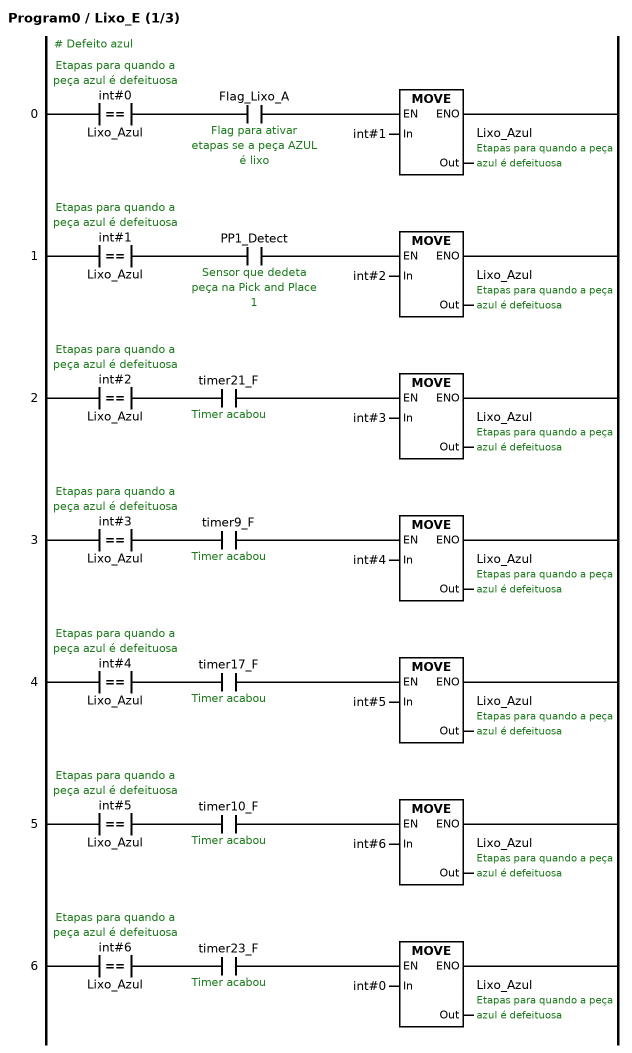
(* [picture p120: Program0 / Lixo_E, rungs 0-6] *)
(* Rung 0: # Defeito azul *)
IF (int#0 = Lixo_Azul) AND Flag_Lixo_A THEN Lixo_Azul := int#1; END_IF;
(* Rung 1 *)
IF (int#1 = Lixo_Azul) AND PP1_Detect THEN Lixo_Azul := int#2; END_IF;
(* Rung 2 *)
IF (int#2 = Lixo_Azul) AND timer21_F THEN Lixo_Azul := int#3; END_IF;
(* Rung 3 *)
IF (int#3 = Lixo_Azul) AND timer9_F THEN Lixo_Azul := int#4; END_IF;
(* Rung 4 *)
IF (int#4 = Lixo_Azul) AND timer17_F THEN Lixo_Azul := int#5; END_IF;
(* Rung 5 *)
IF (int#5 = Lixo_Azul) AND timer10_F THEN Lixo_Azul := int#6; END_IF;
(* Rung 6 *)
IF (int#6 = Lixo_Azul) AND timer23_F THEN Lixo_Azul := int#0; END_IF;

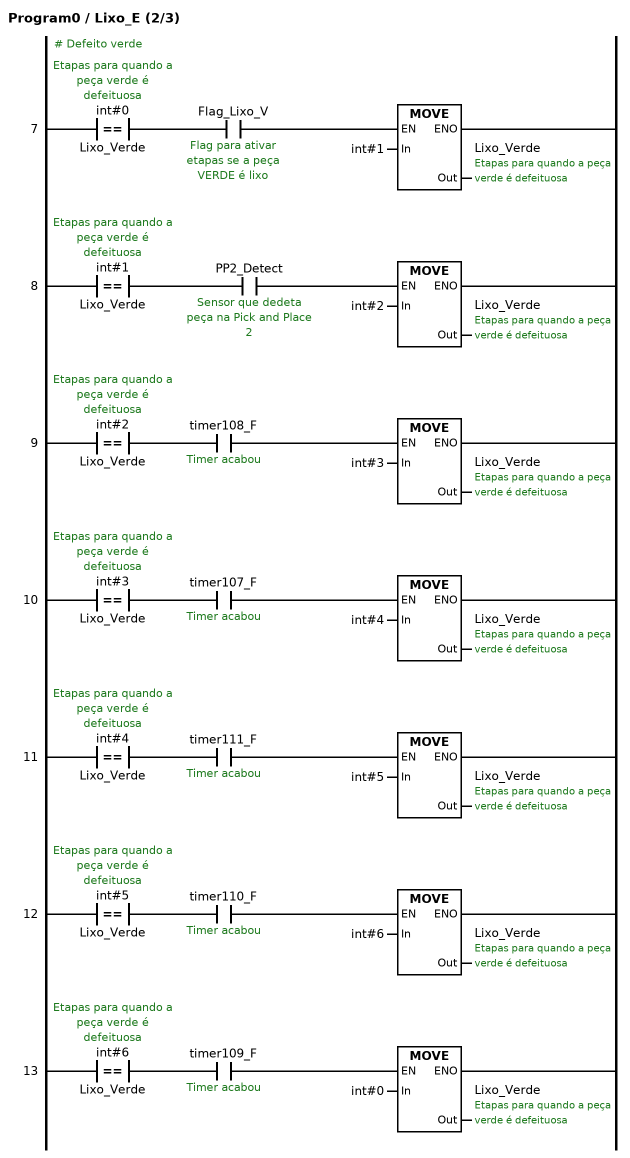
(* Rung 7: # Defeito verde *)
IF (int#0 = Lixo_Verde) AND Flag_Lixo_V THEN Lixo_Verde := int#1; END_IF;
(* Rung 8 *)
IF (int#1 = Lixo_Verde) AND PP2_Detect THEN Lixo_Verde := int#2; END_IF;
(* Rung 9 *)
IF (int#2 = Lixo_Verde) AND timer108_F THEN Lixo_Verde := int#3; END_IF;
(* Rung 10 *)
IF (int#3 = Lixo_Verde) AND timer107_F THEN Lixo_Verde := int#4; END_IF;
(* Rung 11 *)
IF (int#4 = Lixo_Verde) AND timer111_F THEN Lixo_Verde := int#5; END_IF;
(* Rung 12 *)
IF (int#5 = Lixo_Verde) AND timer110_F THEN Lixo_Verde := int#6; END_IF;
(* Rung 13 *)
IF (int#6 = Lixo_Verde) AND timer109_F THEN Lixo_Verde := int#0; END_IF;

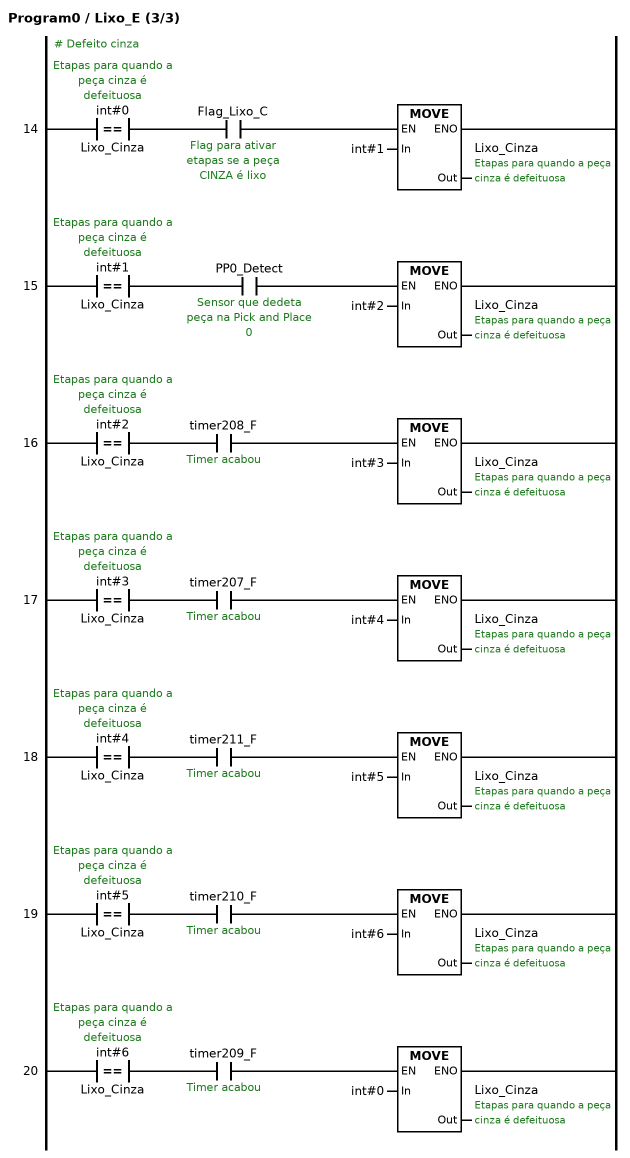
(* Rung 14: # Defeito cinza *)
IF (int#0 = Lixo_Cinza) AND Flag_Lixo_C THEN Lixo_Cinza := int#1; END_IF;
(* Rung 15 *)
IF (int#1 = Lixo_Cinza) AND PP0_Detect THEN Lixo_Cinza := int#2; END_IF;
(* Rung 16 *)
IF (int#2 = Lixo_Cinza) AND timer208_F THEN Lixo_Cinza := int#3; END_IF;
(* Rung 17 *)
IF (int#3 = Lixo_Cinza) AND timer207_F THEN Lixo_Cinza := int#4; END_IF;
(* Rung 18 *)
IF (int#4 = Lixo_Cinza) AND timer211_F THEN Lixo_Cinza := int#5; END_IF;
(* Rung 19 *)
IF (int#5 = Lixo_Cinza) AND timer210_F THEN Lixo_Cinza := int#6; END_IF;
(* Rung 20 *)
IF (int#6 = Lixo_Cinza) AND timer209_F THEN Lixo_Cinza := int#0; END_IF;

(* Section Lixo_S: ladder, written here as Structured Text *)

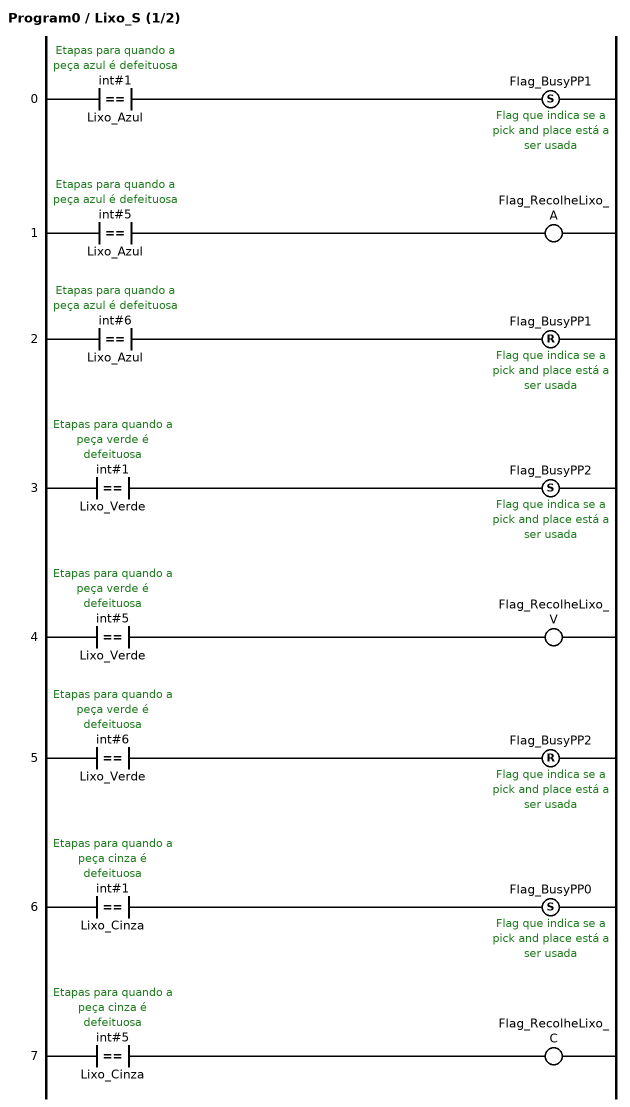
(* Rung 0 *)
IF int#1 = Lixo_Azul THEN Flag_BusyPP1 := TRUE; END_IF;
(* Rung 1 *)
Flag_RecolheLixo_A := int#5 = Lixo_Azul;
(* Rung 2 *)
IF int#6 = Lixo_Azul THEN Flag_BusyPP1 := FALSE; END_IF;
(* Rung 3 *)
IF int#1 = Lixo_Verde THEN Flag_BusyPP2 := TRUE; END_IF;
(* Rung 4 *)
Flag_RecolheLixo_V := int#5 = Lixo_Verde;
(* Rung 5 *)
IF int#6 = Lixo_Verde THEN Flag_BusyPP2 := FALSE; END_IF;
(* Rung 6 *)
IF int#1 = Lixo_Cinza THEN Flag_BusyPP0 := TRUE; END_IF;
(* Rung 7 *)
Flag_RecolheLixo_C := int#5 = Lixo_Cinza;

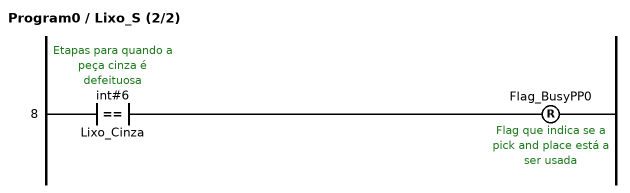
(* Rung 8 *)
IF int#6 = Lixo_Cinza THEN Flag_BusyPP0 := FALSE; END_IF;

(* Section Recolhe_Lixo_E: ladder, written here as Structured Text *)

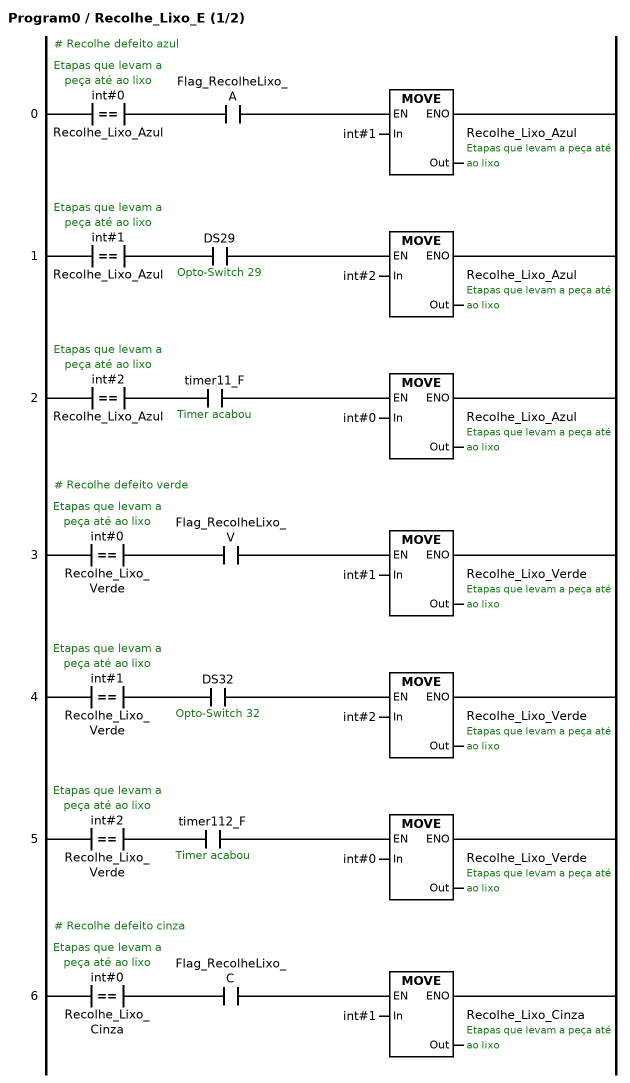
(* Rung 0: # Recolhe defeito azul *)
IF (int#0 = Recolhe_Lixo_Azul) AND Flag_RecolheLixo_A THEN Recolhe_Lixo_Azul := int#1; END_IF;
(* Rung 1 *)
IF (int#1 = Recolhe_Lixo_Azul) AND DS29 THEN Recolhe_Lixo_Azul := int#2; END_IF;
(* Rung 2 *)
IF (int#2 = Recolhe_Lixo_Azul) AND timer11_F THEN Recolhe_Lixo_Azul := int#0; END_IF;
(* Rung 3: # Recolhe defeito verde *)
IF (int#0 = Recolhe_Lixo_Verde) AND Flag_RecolheLixo_V THEN Recolhe_Lixo_Verde := int#1; END_IF;
(* Rung 4 *)
IF (int#1 = Recolhe_Lixo_Verde) AND DS32 THEN Recolhe_Lixo_Verde := int#2; END_IF;
(* Rung 5 *)
IF (int#2 = Recolhe_Lixo_Verde) AND timer112_F THEN Recolhe_Lixo_Verde := int#0; END_IF;
(* Rung 6: # Recolhe defeito cinza *)
IF (int#0 = Recolhe_Lixo_Cinza) AND Flag_RecolheLixo_C THEN Recolhe_Lixo_Cinza := int#1; END_IF;

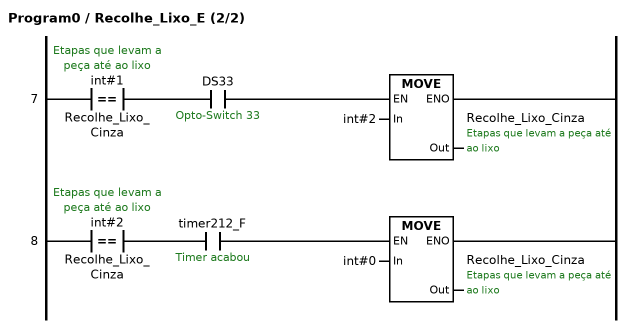
(* Rung 7 *)
IF (int#1 = Recolhe_Lixo_Cinza) AND DS33 THEN Recolhe_Lixo_Cinza := int#2; END_IF;
(* Rung 8 *)
IF (int#2 = Recolhe_Lixo_Cinza) AND timer212_F THEN Recolhe_Lixo_Cinza := int#0; END_IF;

(* Section Recolhe_Lixo_S: ladder, written here as Structured Text *)

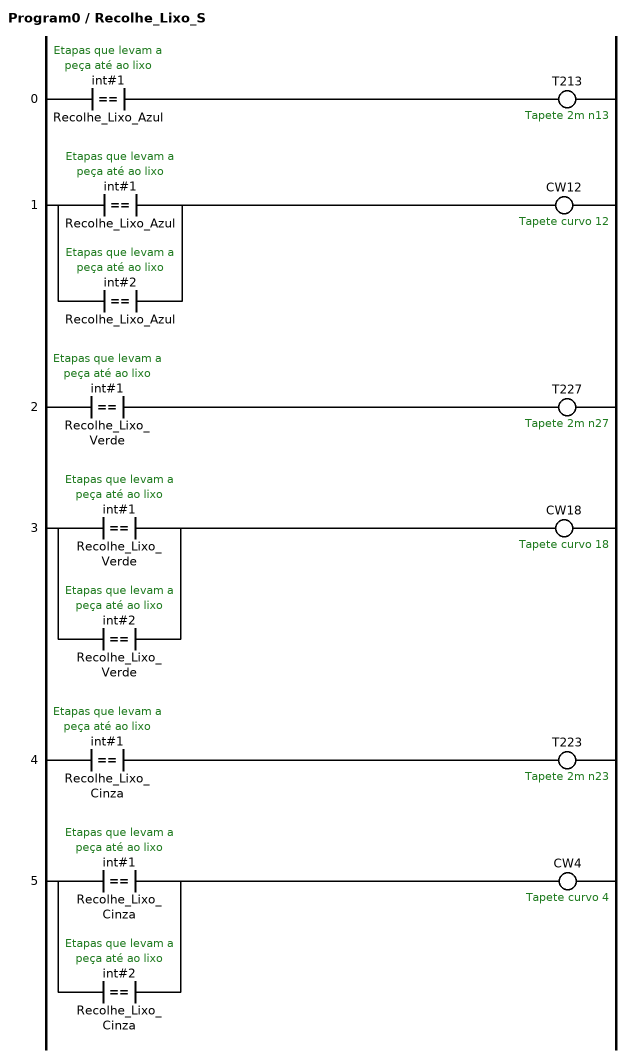
(* Rung 0 *)
T213 := int#1 = Recolhe_Lixo_Azul;
(* Rung 1 *)
CW12 := (int#1 = Recolhe_Lixo_Azul) OR (int#2 = Recolhe_Lixo_Azul);
(* Rung 2 *)
T227 := int#1 = Recolhe_Lixo_Verde;
(* Rung 3 *)
CW18 := (int#1 = Recolhe_Lixo_Verde) OR (int#2 = Recolhe_Lixo_Verde);
(* Rung 4 *)
T223 := int#1 = Recolhe_Lixo_Cinza;
(* Rung 5 *)
CW4 := (int#1 = Recolhe_Lixo_Cinza) OR (int#2 = Recolhe_Lixo_Cinza);

(* Section Repara_Peca_E: ladder, written here as Structured Text *)

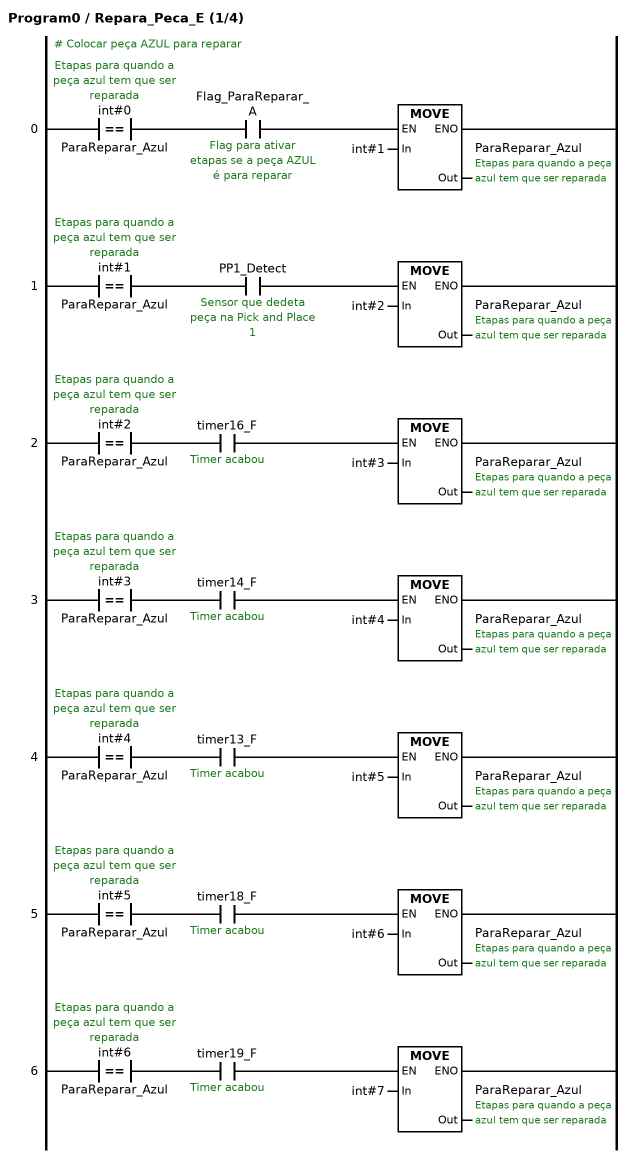
(* Rung 0: # Colocar peça AZUL para reparar *)
IF (int#0 = ParaReparar_Azul) AND Flag_ParaReparar_A THEN ParaReparar_Azul := int#1; END_IF;
(* Rung 1 *)
IF (int#1 = ParaReparar_Azul) AND PP1_Detect THEN ParaReparar_Azul := int#2; END_IF;
(* Rung 2 *)
IF (int#2 = ParaReparar_Azul) AND timer16_F THEN ParaReparar_Azul := int#3; END_IF;
(* Rung 3 *)
IF (int#3 = ParaReparar_Azul) AND timer14_F THEN ParaReparar_Azul := int#4; END_IF;
(* Rung 4 *)
IF (int#4 = ParaReparar_Azul) AND timer13_F THEN ParaReparar_Azul := int#5; END_IF;
(* Rung 5 *)
IF (int#5 = ParaReparar_Azul) AND timer18_F THEN ParaReparar_Azul := int#6; END_IF;
(* Rung 6 *)
IF (int#6 = ParaReparar_Azul) AND timer19_F THEN ParaReparar_Azul := int#7; END_IF;

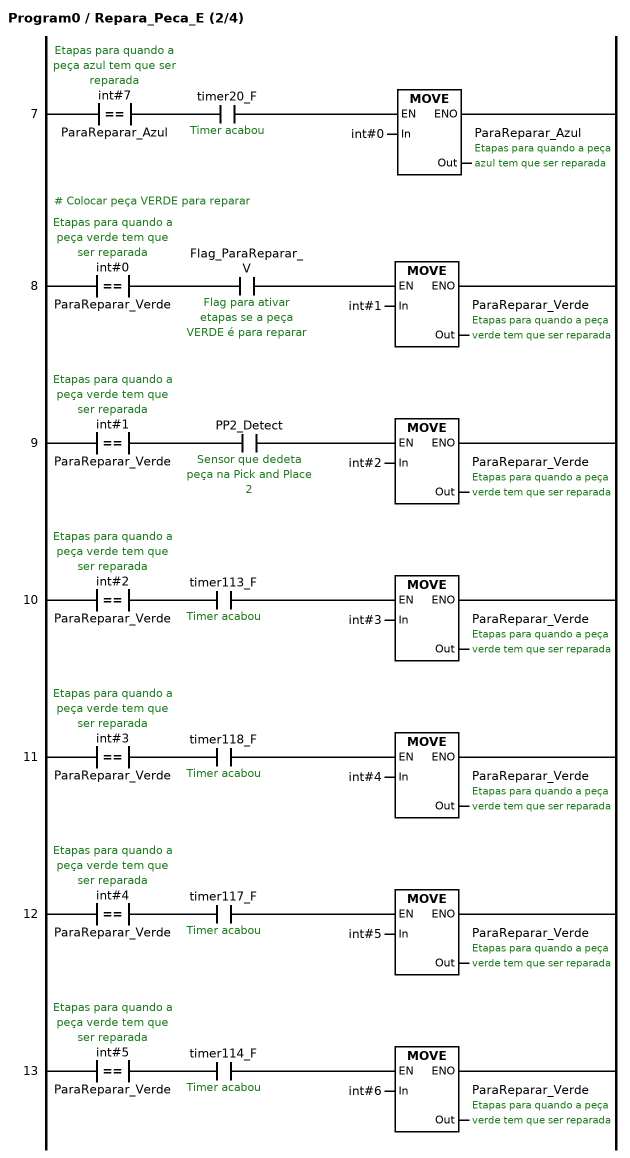
(* Rung 7 *)
IF (int#7 = ParaReparar_Azul) AND timer20_F THEN ParaReparar_Azul := int#0; END_IF;
(* Rung 8: # Colocar peça VERDE para reparar *)
IF (int#0 = ParaReparar_Verde) AND Flag_ParaReparar_V THEN ParaReparar_Verde := int#1; END_IF;
(* Rung 9 *)
IF (int#1 = ParaReparar_Verde) AND PP2_Detect THEN ParaReparar_Verde := int#2; END_IF;
(* Rung 10 *)
IF (int#2 = ParaReparar_Verde) AND timer113_F THEN ParaReparar_Verde := int#3; END_IF;
(* Rung 11 *)
IF (int#3 = ParaReparar_Verde) AND timer118_F THEN ParaReparar_Verde := int#4; END_IF;
(* Rung 12 *)
IF (int#4 = ParaReparar_Verde) AND timer117_F THEN ParaReparar_Verde := int#5; END_IF;
(* Rung 13 *)
IF (int#5 = ParaReparar_Verde) AND timer114_F THEN ParaReparar_Verde := int#6; END_IF;

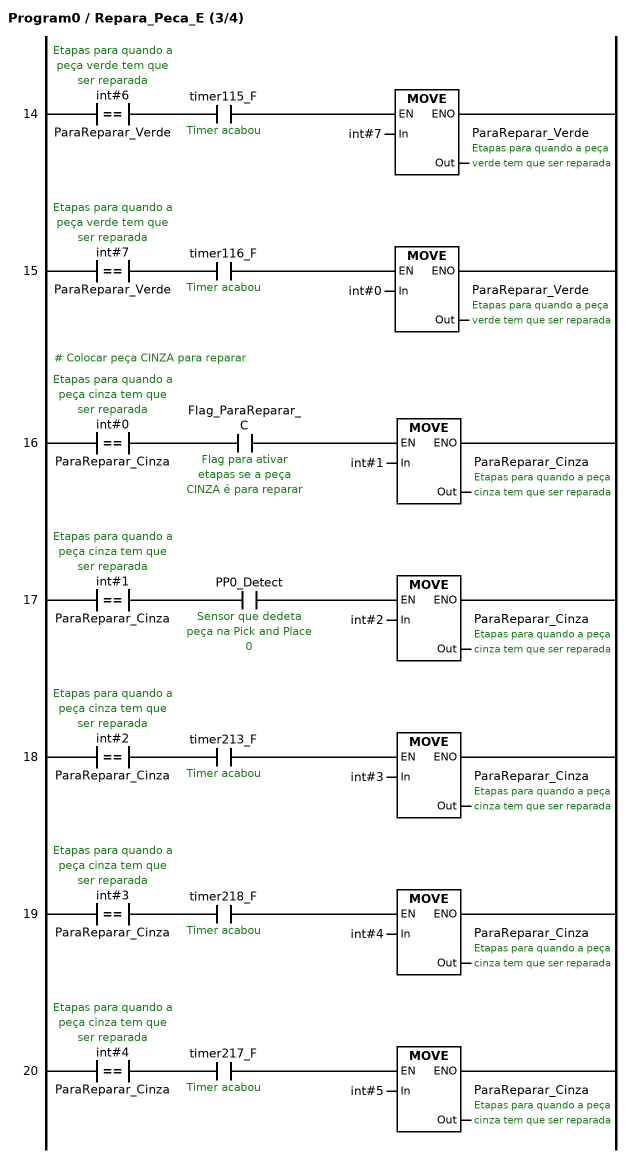
(* Rung 14 *)
IF (int#6 = ParaReparar_Verde) AND timer115_F THEN ParaReparar_Verde := int#7; END_IF;
(* Rung 15 *)
IF (int#7 = ParaReparar_Verde) AND timer116_F THEN ParaReparar_Verde := int#0; END_IF;
(* Rung 16: # Colocar peça CINZA para reparar *)
IF (int#0 = ParaReparar_Cinza) AND Flag_ParaReparar_C THEN ParaReparar_Cinza := int#1; END_IF;
(* Rung 17 *)
IF (int#1 = ParaReparar_Cinza) AND PP0_Detect THEN ParaReparar_Cinza := int#2; END_IF;
(* Rung 18 *)
IF (int#2 = ParaReparar_Cinza) AND timer213_F THEN ParaReparar_Cinza := int#3; END_IF;
(* Rung 19 *)
IF (int#3 = ParaReparar_Cinza) AND timer218_F THEN ParaReparar_Cinza := int#4; END_IF;
(* Rung 20 *)
IF (int#4 = ParaReparar_Cinza) AND timer217_F THEN ParaReparar_Cinza := int#5; END_IF;

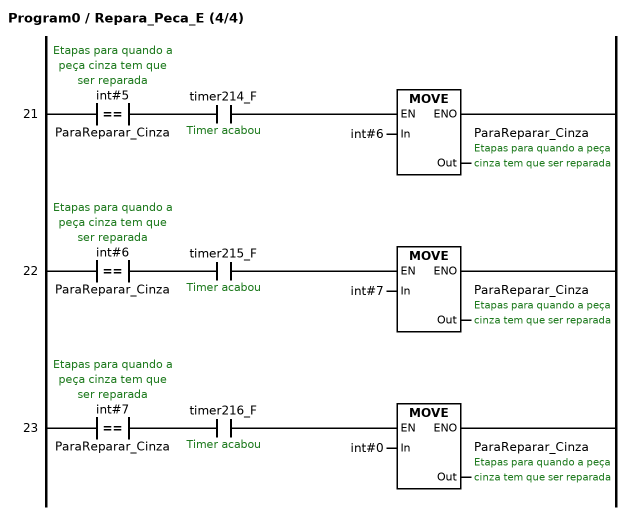
(* Rung 21 *)
IF (int#5 = ParaReparar_Cinza) AND timer214_F THEN ParaReparar_Cinza := int#6; END_IF;
(* Rung 22 *)
IF (int#6 = ParaReparar_Cinza) AND timer215_F THEN ParaReparar_Cinza := int#7; END_IF;
(* Rung 23 *)
IF (int#7 = ParaReparar_Cinza) AND timer216_F THEN ParaReparar_Cinza := int#0; END_IF;

(* Section Repara_Peca_S: ladder, written here as Structured Text *)

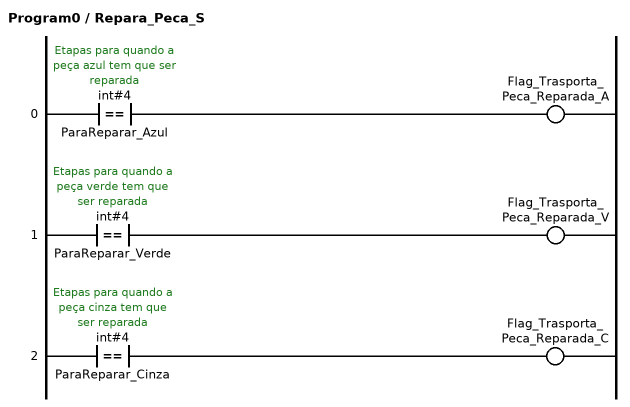
(* Rung 0 *)
Flag_Trasporta_Peca_Reparada_A := int#4 = ParaReparar_Azul;
(* Rung 1 *)
Flag_Trasporta_Peca_Reparada_V := int#4 = ParaReparar_Verde;
(* Rung 2 *)
Flag_Trasporta_Peca_Reparada_C := int#4 = ParaReparar_Cinza;

(* Section Recolhe_PR_E: ladder, written here as Structured Text *)

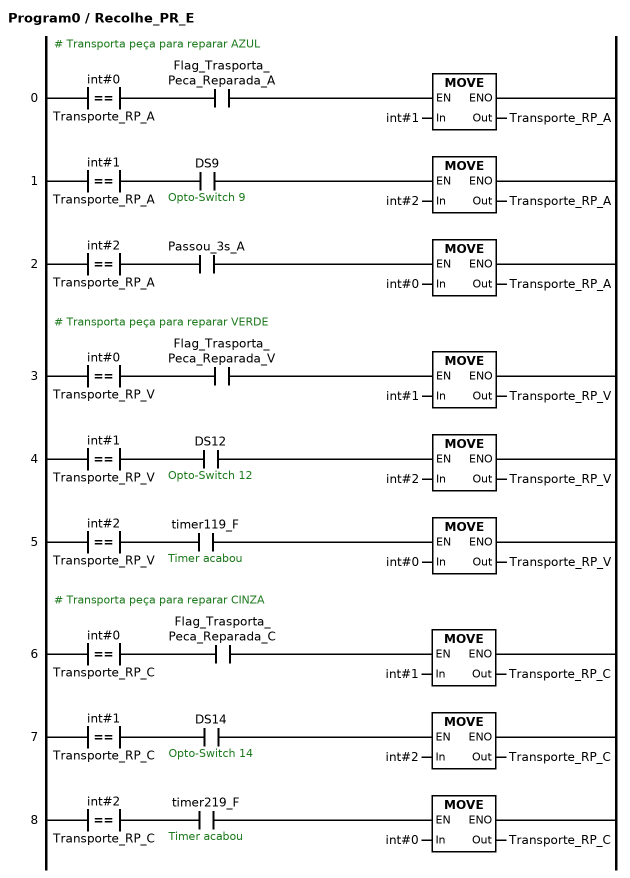
(* Rung 0: # Transporta peça para reparar AZUL *)
IF (int#0 = Transporte_RP_A) AND Flag_Trasporta_Peca_Reparada_A THEN Transporte_RP_A := int#1; END_IF;
(* Rung 1 *)
IF (int#1 = Transporte_RP_A) AND DS9 THEN Transporte_RP_A := int#2; END_IF;
(* Rung 2 *)
IF (int#2 = Transporte_RP_A) AND Passou_3s_A THEN Transporte_RP_A := int#0; END_IF;
(* Rung 3: # Transporta peça para reparar VERDE *)
IF (int#0 = Transporte_RP_V) AND Flag_Trasporta_Peca_Reparada_V THEN Transporte_RP_V := int#1; END_IF;
(* Rung 4 *)
IF (int#1 = Transporte_RP_V) AND DS12 THEN Transporte_RP_V := int#2; END_IF;
(* Rung 5 *)
IF (int#2 = Transporte_RP_V) AND timer119_F THEN Transporte_RP_V := int#0; END_IF;
(* Rung 6: # Transporta peça para reparar CINZA *)
IF (int#0 = Transporte_RP_C) AND Flag_Trasporta_Peca_Reparada_C THEN Transporte_RP_C := int#1; END_IF;
(* Rung 7 *)
IF (int#1 = Transporte_RP_C) AND DS14 THEN Transporte_RP_C := int#2; END_IF;
(* Rung 8 *)
IF (int#2 = Transporte_RP_C) AND timer219_F THEN Transporte_RP_C := int#0; END_IF;

(* Section Recolhe_PR_S: ladder, written here as Structured Text *)

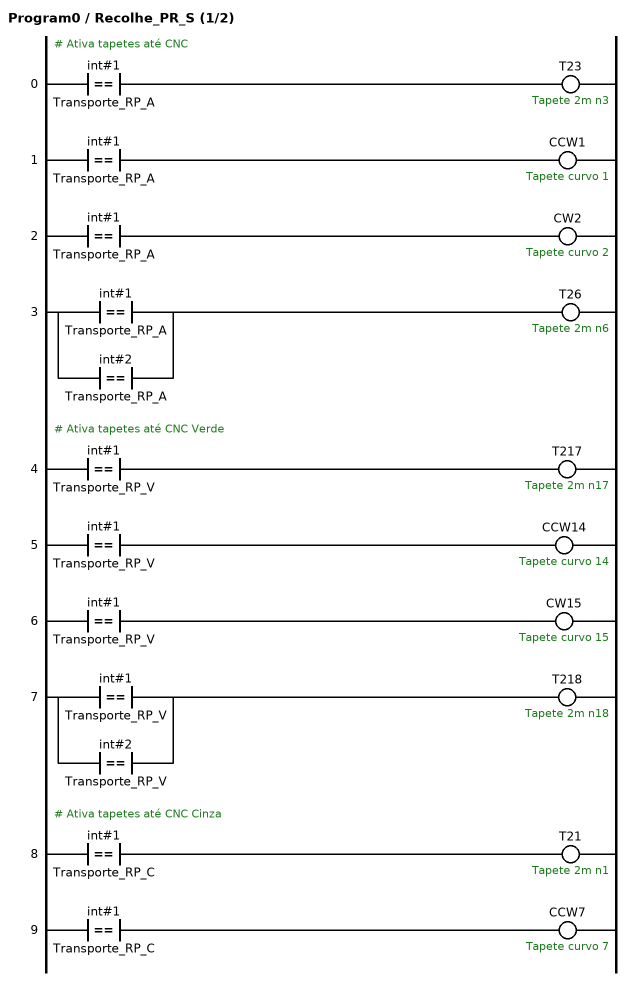
(* Rung 0: # Ativa tapetes até CNC *)
T23 := int#1 = Transporte_RP_A;
(* Rung 1 *)
CCW1 := int#1 = Transporte_RP_A;
(* Rung 2 *)
CW2 := int#1 = Transporte_RP_A;
(* Rung 3 *)
T26 := (int#1 = Transporte_RP_A) OR (int#2 = Transporte_RP_A);
(* Rung 4: # Ativa tapetes até CNC Verde *)
T217 := int#1 = Transporte_RP_V;
(* Rung 5 *)
CCW14 := int#1 = Transporte_RP_V;
(* Rung 6 *)
CW15 := int#1 = Transporte_RP_V;
(* Rung 7 *)
T218 := (int#1 = Transporte_RP_V) OR (int#2 = Transporte_RP_V);
(* Rung 8: # Ativa tapetes até CNC Cinza *)
T21 := int#1 = Transporte_RP_C;
(* Rung 9 *)
CCW7 := int#1 = Transporte_RP_C;

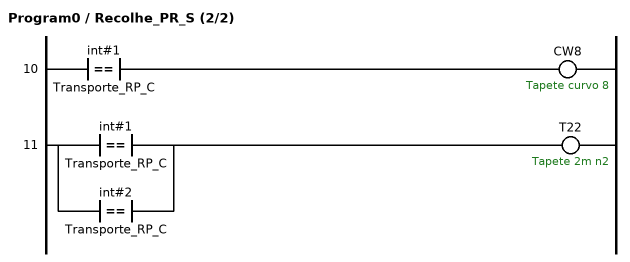
(* Rung 10 *)
CW8 := int#1 = Transporte_RP_C;
(* Rung 11 *)
T22 := (int#1 = Transporte_RP_C) OR (int#2 = Transporte_RP_C);

(* Section Saida_CNC_E: ladder, written here as Structured Text *)

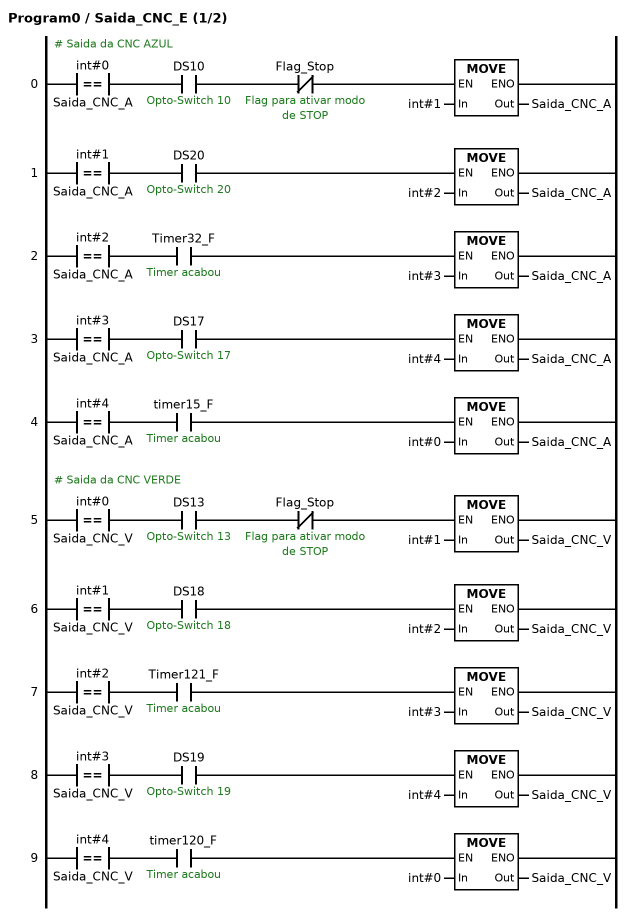
(* Rung 0: # Saida da CNC AZUL *)
IF (int#0 = Saida_CNC_A) AND DS10 AND NOT Flag_Stop THEN Saida_CNC_A := int#1; END_IF;
(* Rung 1 *)
IF (int#1 = Saida_CNC_A) AND DS20 THEN Saida_CNC_A := int#2; END_IF;
(* Rung 2 *)
IF (int#2 = Saida_CNC_A) AND Timer32_F THEN Saida_CNC_A := int#3; END_IF;
(* Rung 3 *)
IF (int#3 = Saida_CNC_A) AND DS17 THEN Saida_CNC_A := int#4; END_IF;
(* Rung 4 *)
IF (int#4 = Saida_CNC_A) AND timer15_F THEN Saida_CNC_A := int#0; END_IF;
(* Rung 5: # Saida da CNC VERDE *)
IF (int#0 = Saida_CNC_V) AND DS13 AND NOT Flag_Stop THEN Saida_CNC_V := int#1; END_IF;
(* Rung 6 *)
IF (int#1 = Saida_CNC_V) AND DS18 THEN Saida_CNC_V := int#2; END_IF;
(* Rung 7 *)
IF (int#2 = Saida_CNC_V) AND Timer121_F THEN Saida_CNC_V := int#3; END_IF;
(* Rung 8 *)
IF (int#3 = Saida_CNC_V) AND DS19 THEN Saida_CNC_V := int#4; END_IF;
(* Rung 9 *)
IF (int#4 = Saida_CNC_V) AND timer120_F THEN Saida_CNC_V := int#0; END_IF;

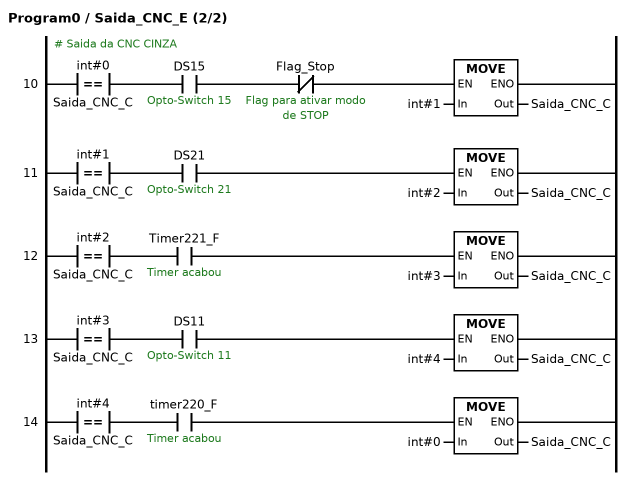
(* Rung 10: # Saida da CNC CINZA *)
IF (int#0 = Saida_CNC_C) AND DS15 AND NOT Flag_Stop THEN Saida_CNC_C := int#1; END_IF;
(* Rung 11 *)
IF (int#1 = Saida_CNC_C) AND DS21 THEN Saida_CNC_C := int#2; END_IF;
(* Rung 12 *)
IF (int#2 = Saida_CNC_C) AND Timer221_F THEN Saida_CNC_C := int#3; END_IF;
(* Rung 13 *)
IF (int#3 = Saida_CNC_C) AND DS11 THEN Saida_CNC_C := int#4; END_IF;
(* Rung 14 *)
IF (int#4 = Saida_CNC_C) AND timer220_F THEN Saida_CNC_C := int#0; END_IF;

(* Section Saida_CNC_S: ladder, written here as Structured Text *)

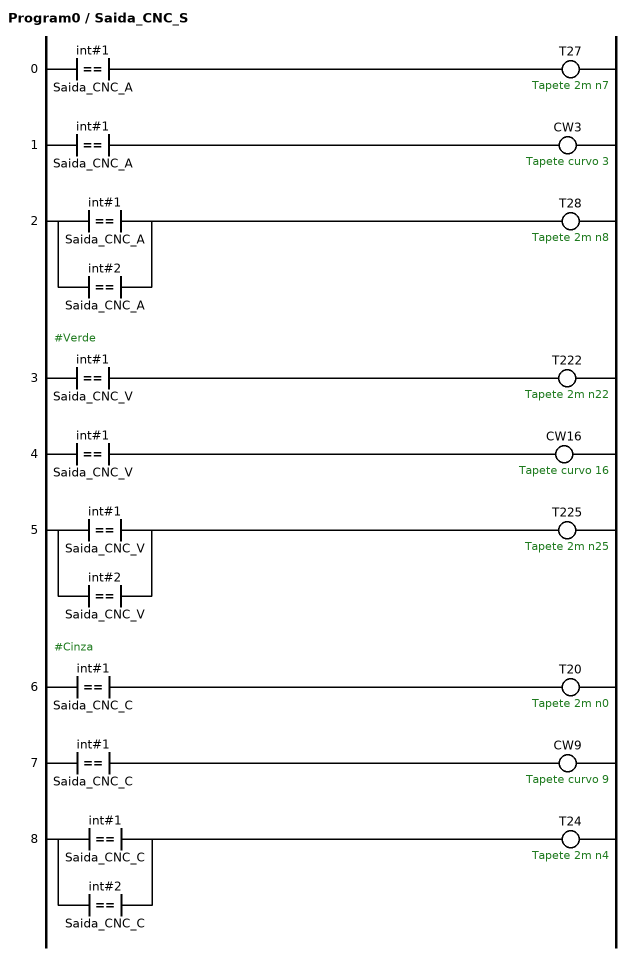
(* Rung 0 *)
T27 := int#1 = Saida_CNC_A;
(* Rung 1 *)
CW3 := int#1 = Saida_CNC_A;
(* Rung 2 *)
T28 := (int#1 = Saida_CNC_A) OR (int#2 = Saida_CNC_A);
(* Rung 3: #Verde *)
T222 := int#1 = Saida_CNC_V;
(* Rung 4 *)
CW16 := int#1 = Saida_CNC_V;
(* Rung 5 *)
T225 := (int#1 = Saida_CNC_V) OR (int#2 = Saida_CNC_V);
(* Rung 6: #Cinza *)
T20 := int#1 = Saida_CNC_C;
(* Rung 7 *)
CW9 := int#1 = Saida_CNC_C;
(* Rung 8 *)
T24 := (int#1 = Saida_CNC_C) OR (int#2 = Saida_CNC_C);

(* Section Stock_E: ladder, written here as Structured Text *)

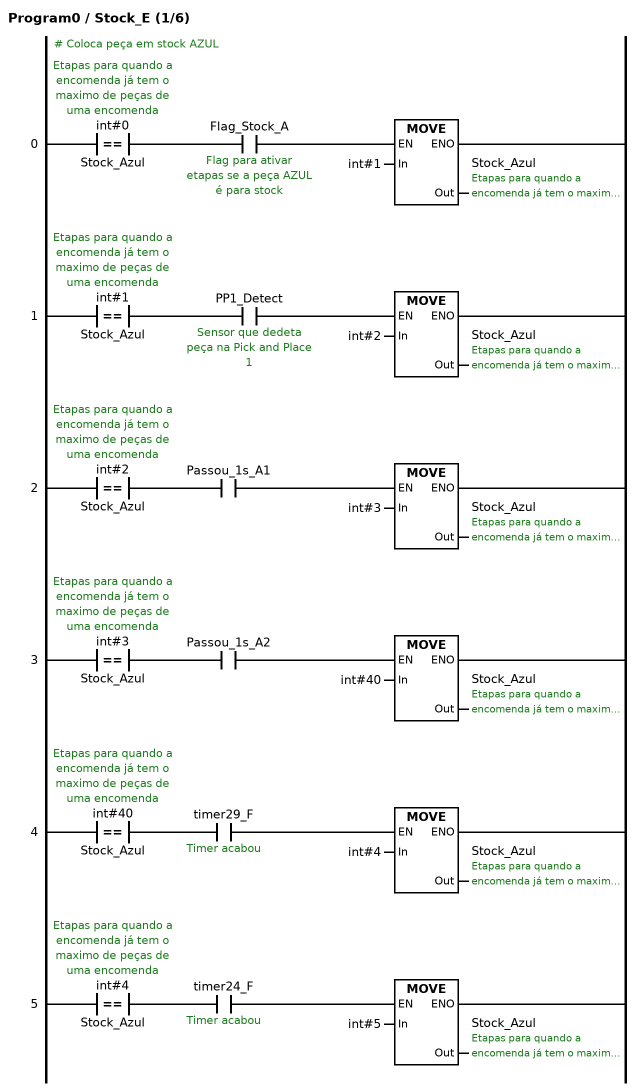
(* Rung 0: # Coloca peça em stock AZUL *)
IF (int#0 = Stock_Azul) AND Flag_Stock_A THEN Stock_Azul := int#1; END_IF;
(* Rung 1 *)
IF (int#1 = Stock_Azul) AND PP1_Detect THEN Stock_Azul := int#2; END_IF;
(* Rung 2 *)
IF (int#2 = Stock_Azul) AND Passou_1s_A1 THEN Stock_Azul := int#3; END_IF;
(* Rung 3 *)
IF (int#3 = Stock_Azul) AND Passou_1s_A2 THEN Stock_Azul := int#40; END_IF;
(* Rung 4 *)
IF (int#40 = Stock_Azul) AND timer29_F THEN Stock_Azul := int#4; END_IF;
(* Rung 5 *)
IF (int#4 = Stock_Azul) AND timer24_F THEN Stock_Azul := int#5; END_IF;

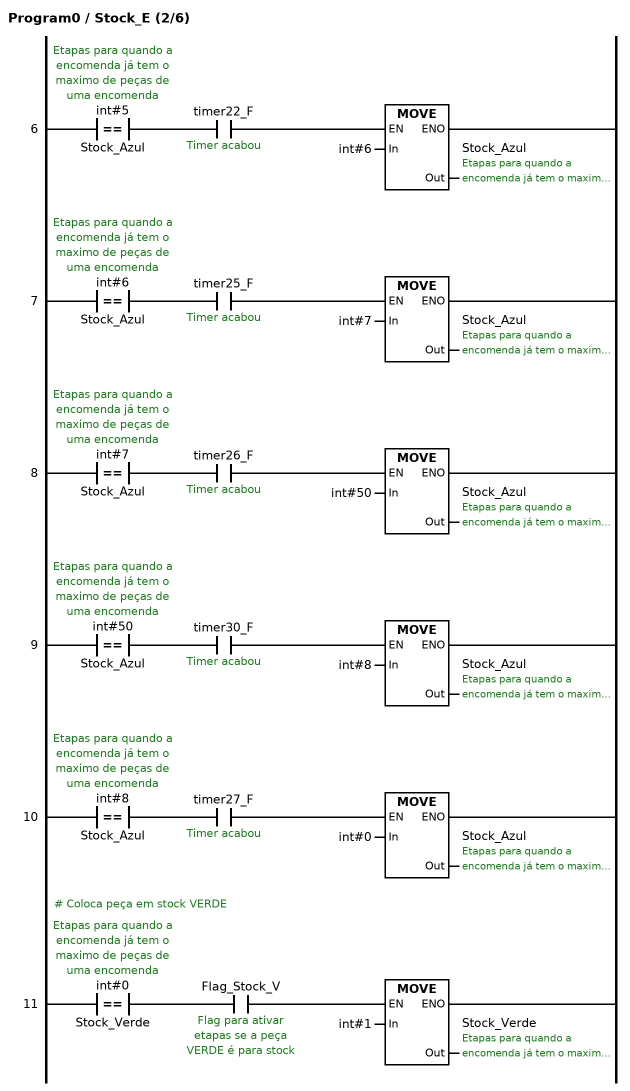
(* Rung 6 *)
IF (int#5 = Stock_Azul) AND timer22_F THEN Stock_Azul := int#6; END_IF;
(* Rung 7 *)
IF (int#6 = Stock_Azul) AND timer25_F THEN Stock_Azul := int#7; END_IF;
(* Rung 8 *)
IF (int#7 = Stock_Azul) AND timer26_F THEN Stock_Azul := int#50; END_IF;
(* Rung 9 *)
IF (int#50 = Stock_Azul) AND timer30_F THEN Stock_Azul := int#8; END_IF;
(* Rung 10 *)
IF (int#8 = Stock_Azul) AND timer27_F THEN Stock_Azul := int#0; END_IF;
(* Rung 11: # Coloca peça em stock VERDE *)
IF (int#0 = Stock_Verde) AND Flag_Stock_V THEN Stock_Verde := int#1; END_IF;

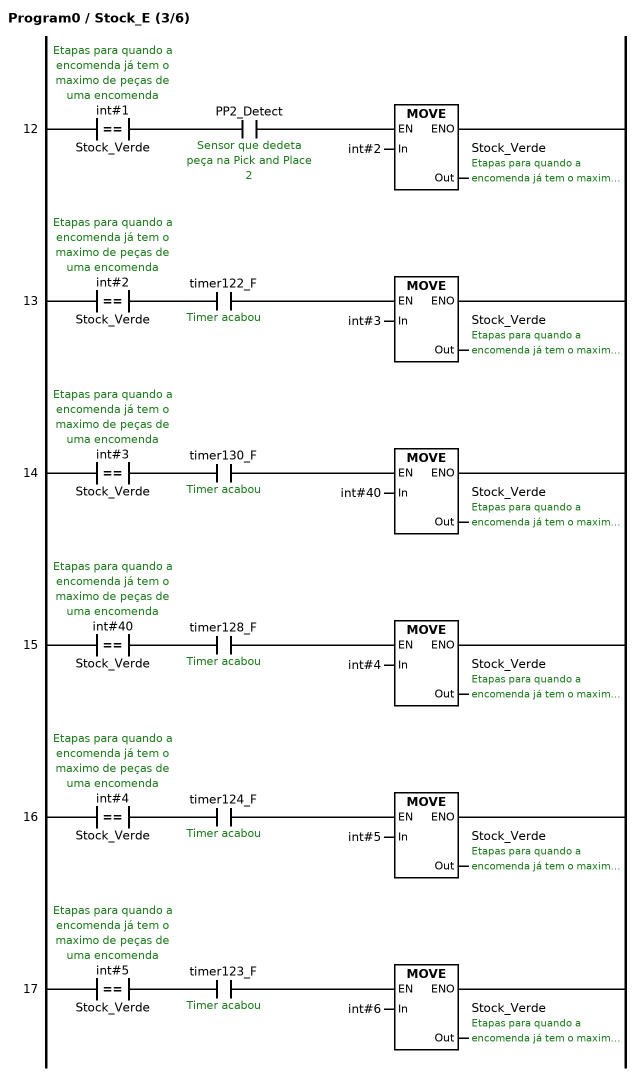
(* Rung 12 *)
IF (int#1 = Stock_Verde) AND PP2_Detect THEN Stock_Verde := int#2; END_IF;
(* Rung 13 *)
IF (int#2 = Stock_Verde) AND timer122_F THEN Stock_Verde := int#3; END_IF;
(* Rung 14 *)
IF (int#3 = Stock_Verde) AND timer130_F THEN Stock_Verde := int#40; END_IF;
(* Rung 15 *)
IF (int#40 = Stock_Verde) AND timer128_F THEN Stock_Verde := int#4; END_IF;
(* Rung 16 *)
IF (int#4 = Stock_Verde) AND timer124_F THEN Stock_Verde := int#5; END_IF;
(* Rung 17 *)
IF (int#5 = Stock_Verde) AND timer123_F THEN Stock_Verde := int#6; END_IF;

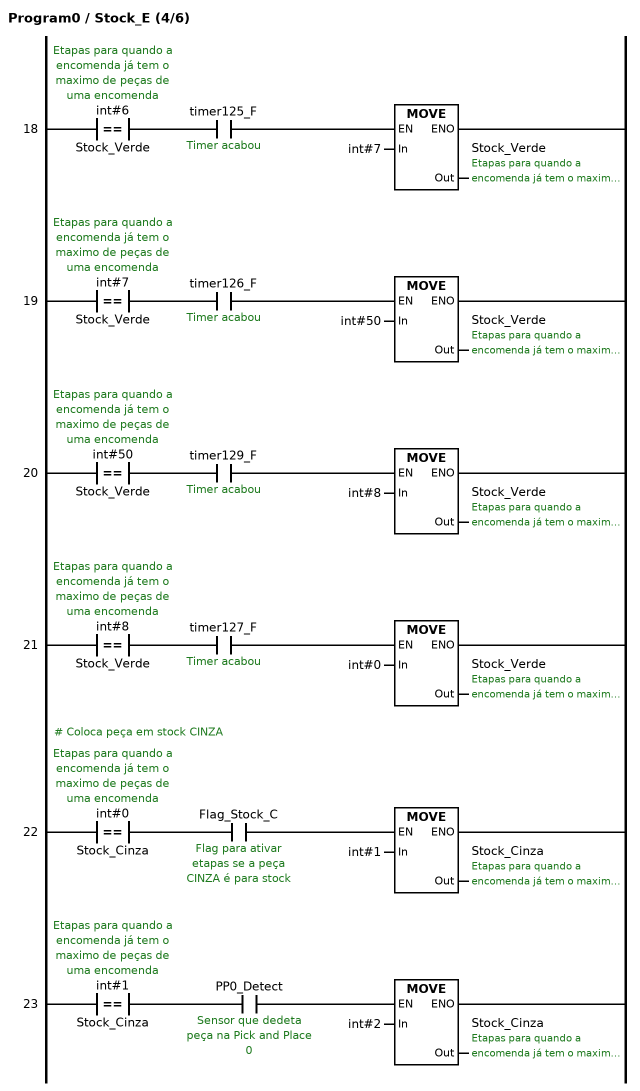
(* Rung 18 *)
IF (int#6 = Stock_Verde) AND timer125_F THEN Stock_Verde := int#7; END_IF;
(* Rung 19 *)
IF (int#7 = Stock_Verde) AND timer126_F THEN Stock_Verde := int#50; END_IF;
(* Rung 20 *)
IF (int#50 = Stock_Verde) AND timer129_F THEN Stock_Verde := int#8; END_IF;
(* Rung 21 *)
IF (int#8 = Stock_Verde) AND timer127_F THEN Stock_Verde := int#0; END_IF;
(* Rung 22: # Coloca peça em stock CINZA *)
IF (int#0 = Stock_Cinza) AND Flag_Stock_C THEN Stock_Cinza := int#1; END_IF;
(* Rung 23 *)
IF (int#1 = Stock_Cinza) AND PP0_Detect THEN Stock_Cinza := int#2; END_IF;

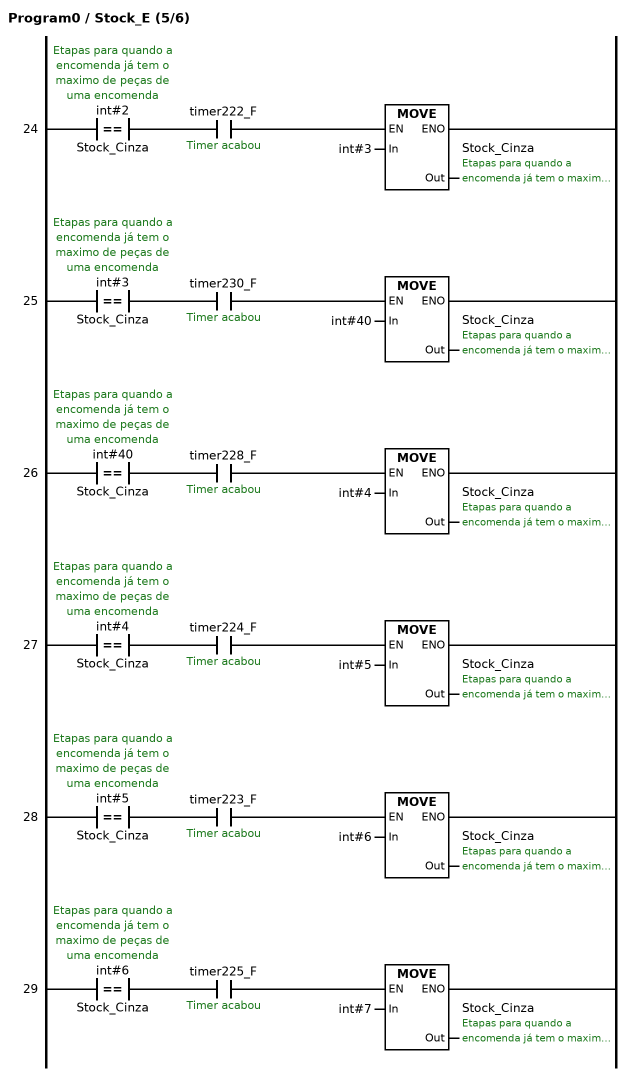
(* Rung 24 *)
IF (int#2 = Stock_Cinza) AND timer222_F THEN Stock_Cinza := int#3; END_IF;
(* Rung 25 *)
IF (int#3 = Stock_Cinza) AND timer230_F THEN Stock_Cinza := int#40; END_IF;
(* Rung 26 *)
IF (int#40 = Stock_Cinza) AND timer228_F THEN Stock_Cinza := int#4; END_IF;
(* Rung 27 *)
IF (int#4 = Stock_Cinza) AND timer224_F THEN Stock_Cinza := int#5; END_IF;
(* Rung 28 *)
IF (int#5 = Stock_Cinza) AND timer223_F THEN Stock_Cinza := int#6; END_IF;
(* Rung 29 *)
IF (int#6 = Stock_Cinza) AND timer225_F THEN Stock_Cinza := int#7; END_IF;

